Staubli VAL3: CalAdjustZ.pgx

public program CalAdjustZ()
  local num l_nDistance
  local trsf l_trZ
  local num l_nDir
begin
  l_nDistance=distance(db:pAdjustZ_2_1,db:pAdjustZ_2_2)
  switch db:sMounting
    case "Floor"
      l_nDir=1
    break
    case "Ceiling"
      l_nDir=-1
    break
    default
      l_nDir=1
    break
  endSwitch
  //
  if db:pAdjustZ_2_1.trsf.z<db:pAdjustZ_2_2.trsf.z
    l_trZ={0,0,-l_nDistance*l_nDir,0,0,0}
  else
    l_trZ={0,0,l_nDistance*l_nDir,0,0,0}
  endIf
  //
  db:tTool3.trsf=db:utCurrentTool.tValue.trsf*l_trZ
  db:tTool3.trsf.rx=db:tTool1.trsf.rx
  db:tTool3.trsf.ry=db:tTool1.trsf.ry
  db:tTool3.trsf.rz=db:tTool1.trsf.rz
  call db:hmiAlert("SaveInTool3","info")
end
